// Mitsubishi GX Works2 project: 두번째시간   PLC: Q02/Q02H

PROGRAM MAIN
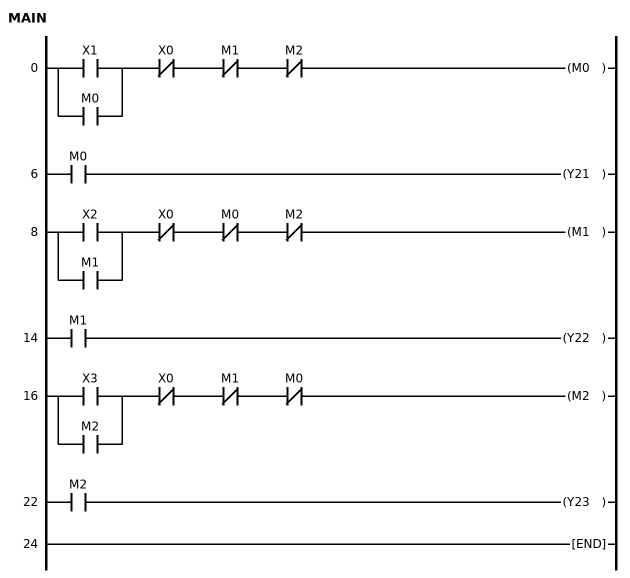
0     LD      X1
      OR      M0
      ANI     X0
      ANI     M1
      ANI     M2
      OUT     M0
6     LD      M0
      OUT     Y21
8     LD      X2
      OR      M1
      ANI     X0
      ANI     M0
      ANI     M2
      OUT     M1
14    LD      M1
      OUT     Y22
16    LD      X3
      OR      M2
      ANI     X0
      ANI     M1
      ANI     M0
      OUT     M2
22    LD      M2
      OUT     Y23
24    END
END_PROGRAM
